# EPICS substitutions: examples/PSI/plugins/cpp_logic/examples/cpp_logic_waveform/cfg/libmain.so_cpp_logic.subs
# Auto-generated C++ logic substitutions
# Logic: cpp_logic_waveform

file ecmcCppLogicWaveformIn.template {
  pattern { REC, PARAM, DESC, NELM, FTVL, DTYP }
  { "epics-ec-s23-mm-analogOutputArray01", "epics_ec.s23.mm.analogOutputArray01", "epics_ec.s23.mm.analogOutputArray01", "100", "SHORT", "asynInt16ArrayIn" }
}
